(* IEC 61131-3 sources: Caravan/Archiv/12-04-19/Stations/Terminal/HMI/Class/_XMLReader (part 2) *)

  TextLen := _strlen(pText);
  TextLen += 1; // zero termination

  pDest^.pText$^void := StdLib.Malloc(TextLen);
  if pDest^.pText = NIL then
    XmlState := _ERROR;
    retcode := -2;
    return;
  end_if;

  _strcpy(pDest^.pText, pText);

  retcode := 0;

END_FUNCTION //AddTextAscii

FUNCTION _XMLReader::AddTextUni
	VAR_INPUT
		pDest 	: ^_XML_ELEMENT;
		pText 	: ^UINT;
	END_VAR
	VAR_OUTPUT
		retcode 	: DINT;
	END_VAR
  VAR
  	TextLen   : UDINT;
  END_VAR

  retcode := -1;

  if (pDest = NIL) | (pText = NIL) then
    return;
  end_if;

  // only allowed to add text when element has no children or already has a text
  if (pDest^.pText <> NIL) | (pDest^.pChildren <> NIL) then
    return;
  end_if;

  TextLen := SigCLib.StrLen16(pText)*2;
  TextLen += 2; // zero termination

  pDest^.pText$^void := StdLib.Malloc(TextLen);
  if pDest^.pText = NIL then
    XmlState := _ERROR;
    retcode := -2;
    return;
  end_if;

  SigCLib.StrCpy16(pDest^.pText$^UINT, pText);

  retcode := 0;

END_FUNCTION //AddTextUni

FUNCTION _XMLReader::CreateStructAscii
	VAR_INPUT
		parsedBytes 	: ^UDINT;
	END_VAR
	VAR_OUTPUT
		retcode 	: BOOL;
	END_VAR
VAR
	strBuff     : ^USINT;   // first tmp-Buffer
	strBuff2    : ^USINT;   // second tmp-Buffer
  pRun        : ^USINT;   // pointer to go through the information we read
  pStart      : ^USINT;   // points to the start of an element-name, atrib-name, attrib-value and so on...
  signCount   : UDINT;    // counts how much signs a string has
  counter     : UDINT;    // counter how far we passed through the information
  bufferLen   : UDINT;    // size of first buffer
  bufferLen2  : UDINT;    // size of second Buffer
END_VAR

  retcode := FALSE;

  // biggest work will be here
  // we have to go through the buffer and create our XML_STRUCT out of the information
  pRun := pFileBuffer;

  // set start size of buffer to 200, so in most cases we aren't going to resize the buffer
  // (normally names, values aren't this size, maybe text will be longer)
  bufferLen := 200;
  bufferLen2 := 200;

  strBuff$^void := StdLib.Malloc(bufferLen+1);
  strBuff2$^void := StdLib.Malloc(bufferLen2+1);

  if (strBuff = NIL) | (strBuff2 = NIL) then
    XmlState := _ERROR;
    return;
  end_if;

  _memset(strBuff, 0, bufferLen);
  _memset(strBuff2, 0, bufferLen2);

  counter := 1;

  // first handle the header
  if (pRun^ = XML_START) & ((pRun+1)^ = '?') then

    pStart := pRun;
    signCount := 0;

    while pRun^ <> XML_END do
      signCount += 1;

      counter += 1;
      pRun += 1;
    end_while;

    // now we are pointing at the end-mark, this also has to be in the header -> increase counters
    counter += 1;
    signCount += 1;

    if signCount > XML_MAX_HEADER_LENGTH then
      return;
    end_if;

    xmlStruct.Header$^void := StdLib.Malloc(signCount+1);
    _memset(xmlStruct.Header, 0, signCount+1);
    _memcpy(xmlStruct.Header, pStart, signCount);

    // alloc memory for first element and set struct for creator
    xmlStruct.MajorElement$^void := StdLib.Malloc(sizeof(_XML_ELEMENT));
    if (xmlStruct.MajorElement = NIL) then
      XmlState := _ERROR;
      return;
    end_if;
    _memset(xmlStruct.MajorElement, 0, sizeof(_XML_ELEMENT));
    StructCreator.SetStructPtr(#xmlStruct);

  else
    // xml does not start with the header
    ErrorState := _PARSE_ERR_NO_HEADER;
    parsedBytes^ := counter;
    return;
  end_if;

  // now lets see if we find a CR or LF and no signs between except of SPACE
  counter += 1;
  pRun += 1;
  while (pRun^ <> XML_CR) & (pRun^ <> XML_LF) do

    if pRun^ <> XML_SPACE then
      ErrorState := _PARSE_ERR_UNEXPECTED_SIGN;
      parsedBytes^ := counter;
      return; //wrong sign
    end_if;

    counter += 1;
    pRun += 1;
  end_while;

  // Header finished -> now lets start with looking for an Element
  searchFor := _SEARCH_ELEMENT;

  while counter < fileLength do

    case searchFor of

    	_SEARCH_ELEMENT:
    	  // look for '<'
        while pRun^ <> XML_START do

          if (pRun^ <> XML_CR) & (pRun^ <> XML_LF) & (pRun^ <> XML_SPACE) & (pRun^ <> XML_TABULATOR) then
            ErrorState := _PARSE_ERR_UNEXPECTED_SIGN;
            parsedBytes^ := counter;
            return; //wrong sign
          end_if;

          pRun += 1;
          counter += 1;
        end_while;

        // now we are pointing at start-mark, but we need one increase more
        pRun += 1;
        counter += 1;

        if (pRun^ <> XML_SLASH) & (pRun^ <> XML_EXCLAMATION) then
          //START Element
          if bTextSearched = TRUE then
            ErrorState := _PARSE_ERR_UNEXPECTED_SIGN;
            parsedBytes^ := counter;
            return; //wrong sign
          end_if;

          pStart := pRun;
          signCount := 0;

          // next step is to look for Space or End-Mark
          // counter are always one behind the pointer so we do not need to decrease afterwards
          while (pRun^ <> XML_END) & (pRun^ <> XML_SPACE) & (pRun^ <> XML_SLASH) do
            signCount += 1;

            counter += 1;
            pRun += 1;
          end_while;

          // at this point we found an element and we can get the name, so kick off name and add element to struct
          if signCount > bufferLen then
            bufferLen := signCount;
            StdLib.Free(strBuff);

            strBuff$^void := StdLib.Malloc(bufferLen+1);

            if (strBuff = NIL) then
              XmlState := _ERROR;
              return;
            end_if;

          end_if;

          _memcpy(strBuff, pStart, signCount);
          (strBuff+signCount)^ := 0;

          StructCreator.AddElement(strBuff, FALSE);

          // lets see what we have to do next
          if pRun^ = XML_END then

            pRun += 1;
            counter += 1;

            if (pRun^ = XML_CR) | (pRun^ = XML_LF) | (pRun^ = XML_START) | (pRun^ = XML_SPACE) then
              searchFor := _SEARCH_ELEMENT;
            else
              searchFor := _SEARCH_TEXT;
            end_if;

          elsif pRun^ = XML_SLASH then
            StructCreator.CloseElement(NIL,FALSE);

            // element is closed directly -> check if next sign is END-Tag
            pRun += 1;
            counter += 1;

            if pRun^ <> XML_END then
              // no end-tag after slash -> error
              ErrorState := _PARSE_ERR_UNEXPECTED_SIGN;
              parsedBytes^ := counter;
              return; //wrong sign
            end_if;

            // set to next sign
            pRun += 1;
            counter += 1;

            searchFor := _SEARCH_ELEMENT;

          elsif pRun^ = XML_SPACE then
            // in this case there can also be a closing-tag if element ist closed directly
            if (pRun+1)^ = XML_SLASH then

              StructCreator.CloseElement(NIL, FALSE);

              //                      <Element />
              //we point now to the space-----^---
              //but we need to be after end------^
              //this means +3 signs
              pRun += 3;
              counter += 3;

              searchFor := _SEARCH_ELEMENT;
            else
              searchFor := _SEARCH_ATTRIB;
            end_if;

          end_if;

        else
          if pRun^ = XML_SLASH then

            bTextSearched := FALSE;
            // CLOSE Element
            // so just go to the end of the close-element-tag and then close
            pRun += 1;
            counter += 1;

            pStart := pRun;
            signCount := 0;

            while pRun^ <> XML_END do
              signCount += 1;

              counter += 1;
              pRun += 1;
            end_while;

            if signCount > bufferLen then
              bufferLen := signCount;
              StdLib.Free(strBuff);

              strBuff$^void := StdLib.Malloc(bufferLen+1);
              if (strBuff = NIL) then
                XmlState := _ERROR;
                return;
              end_if;
            end_if;

            _memcpy(strBuff, pStart, signCount);
            (strBuff+signCount)^ := 0;

            pRun += 1;
            counter += 1;

            retClose := StructCreator.CloseElement(strBuff, FALSE);
            if retClose <> 0 then
              ErrorState := _PARSE_ERR_WRONG_SEQUENCE;
              parsedBytes^ := counter - signCount - 1;
              return; //wrong sequence of elements
            end_if;

            searchFor := _SEARCH_ELEMENT;

          else
            // check 4 comment
            if bTextSearched = TRUE then
              ErrorState := _PARSE_ERR_UNEXPECTED_SIGN;
              parsedBytes^ := counter;
              return; //wrong sign
            end_if;

            pRun += 1;
            counter += 1;
            if (pRun^ = XML_HYPHEN) & ((pRun+1)^ = XML_HYPHEN) then
              // we found '<!--' this means comment -> skip
              pRun += 2;
              counter += 2;

              while (pRun^ <> XML_HYPHEN) & ((pRun+1)^ <> XML_HYPHEN) & ((pRun+2)^ <> XML_END) do

                pRun += 1;
                counter += 1;

              end_while;
              pRun += 3; // set ptr to one ofter end-tag
              counter += 3;
              // we found the end '-->'
              // go on with searching for an element
              searchFor := _SEARCH_ELEMENT;

            end_if;

          end_if;

        end_if;

      _SEARCH_ATTRIB:

        bTextSearched := FALSE;
    	  // when we have to search 4 an attribute we know that pRun points to a Space
        // so the next sign is the start
        pRun += 1;
        counter += 1;

        pStart := pRun;
        signCount := 0;

        while pRun^ <> XML_EQUAL do

          if (pRun^ = XML_SPACE) | (pRun^ = XML_LF) | (pRun^ = XML_CR) then
            ErrorState := _PARSE_ERR_UNEXPECTED_SIGN;
            parsedBytes^ := counter;
            return; //wrong sign
          end_if;

          signCount += 1;
          counter += 1;
          pRun += 1;
        end_while;

        if signCount > bufferLen then
          bufferLen := signCount;
          StdLib.Free(strBuff);

          strBuff$^void := StdLib.Malloc(bufferLen+1);

          if (strBuff = NIL) then
            XmlState := _ERROR;
            return;
          end_if;

        end_if;

        _memcpy(strBuff, pStart, signCount);
        (strBuff+signCount)^ := 0;

        // we got the name of the attribute now lets get the value

        if ((pRun+1)^ <> XML_QUOTMARK) & ((pRun+1)^ <> XML_APOSTROPHE) then
          ErrorState := _PARSE_ERR_UNEXPECTED_SIGN;
          parsedBytes^ := counter;
          return; // wrong sign
        end_if;

        if ((pRun+1)^ = XML_QUOTMARK) then
          bQuot := TRUE;
        else
          bQuot := FALSE;
        end_if;

        pRun += 2; // set to one after quotation-mark
        counter += 2;

        pStart := pRun;
        signCount := 0;

        while ((pRun^ <> XML_QUOTMARK) & (bQuot = TRUE)) | ((pRun^ <> XML_APOSTROPHE) & (bQuot = FALSE)) do
          signCount += 1;

          counter += 1;
          pRun += 1;
        end_while;

        if signCount > bufferLen2 then
          bufferLen2 := signCount;
          StdLib.Free(strBuff2);

          strBuff2$^void := StdLib.Malloc(bufferLen2+1);

          if (strBuff2 = NIL) then
            XmlState := _ERROR;
            return;
          end_if;

        end_if;

        _memcpy(strBuff2, pStart, signCount);
        (strBuff2+signCount)^ := 0;

        if StructCreator.AddAttribute(strBuff, strBuff2, FALSE) = -1 then
          ErrorState := _PARSE_ERR_ATTRIBUTE_TWICE;
          parsedBytes^ := counter - signCount - 1;
          return; // attribute already exists
        end_if;

        // lets see what we have to do next
        pRun += 1;
        counter += 1;

        if pRun^ = XML_END then
          // so in this case we can have Text afterwards or next thing is an element
          pRun += 1;
          counter += 1;

          if (pRun^ = XML_CR) | (pRun^ = XML_LF) | (pRun^ = XML_START) then
            searchFor := _SEARCH_ELEMENT;
          else
            searchFor := _SEARCH_TEXT;
          end_if;

        elsif pRun^ = XML_SLASH then
            StructCreator.CloseElement(NIL, FALSE);

            // jump one sign after "/>"
            pRun += 2;
            counter += 2;
            searchFor := _SEARCH_ELEMENT;

        elsif pRun^ = XML_SPACE then
          // another attribute
          searchFor := _SEARCH_ATTRIB;
        end_if;

      _SEARCH_TEXT:
        // we already point to the start of the text
        pStart := pRun;
        signCount := 0;

        while pRun^ <> XML_START do
          signCount += 1;

          counter += 1;
          pRun += 1;
        end_while;

        if signCount > bufferLen then
          bufferLen := signCount;
          StdLib.Free(strBuff);

          strBuff$^void := StdLib.Malloc(bufferLen+1);

          if (strBuff = NIL) then
            XmlState := _ERROR;
            return;
          end_if;
        end_if;

        // kick off text & add to actual element
        _memcpy(strBuff, pStart, signCount);
        (strBuff+signCount)^ := 0;

        StructCreator.AddText(strBuff, FALSE);

        //next step hast to be looking for an element
        bTextSearched := TRUE;
        searchFor := _SEARCH_ELEMENT;

    end_case;

  end_while;

  StdLib.Free(strBuff);
  StdLib.Free(strBuff2);

  retcode := TRUE;

END_FUNCTION //CreateStructAscii

FUNCTION _XMLReader::CreateStructUni
	VAR_INPUT
		parsedBytes 	: ^UDINT;
	END_VAR
	VAR_OUTPUT
		retcode 	: BOOL;
	END_VAR
  VAR
    strBuff     : ^USINT;   // first tmp-Buffer
    strBuff2    : ^USINT;   // second tmp-Buffer
    pRun        : ^USINT;   // pointer to go through the information we read
    pStart      : ^USINT;   // points to the start of an element-name, atrib-name, attrib-value and so on...
    signCount   : UDINT;    // counts how much signs a string has
    counter     : UDINT;    // counter how far we passed through the information
    bufferLen   : UDINT;    // size of first buffer
    bufferLen2  : UDINT;    // size of second Buffer
  END_VAR

  retcode := FALSE;

  // biggest work will be here
  // we have to go through the buffer and create our XML_STRUCT out of the information
  pRun := pFileBuffer + 2;

  // set start size of buffer to 200, so in most cases we aren't going to resize the buffer
  // (normally names, values aren't this size, maybe text will be longer)
  bufferLen := 200;
  bufferLen2 := 200;

  strBuff$^void := StdLib.Malloc(bufferLen+2);
  strBuff2$^void := StdLib.Malloc(bufferLen2+2);

  if (strBuff = NIL) | (strBuff2 = NIL) then
    XmlState := _ERROR;
    return;
  end_if;

  _memset(strBuff, 0, bufferLen);
  _memset(strBuff2, 0, bufferLen2);

  counter := 2;

  // first handle the header
  if (pRun^$UINT = XML_START_UNI) & ((pRun+2)^$UINT = 16#003F) then

    pStart := pRun;
    signCount := 0;

    while pRun^$UINT <> XML_END_UNI do
      signCount += 2;

      counter += 2;
      pRun += 2;
    end_while;

    // now we are pointing at the end-mark, this also has to be in the header -> increase counters
    counter += 2;
    signCount += 2;

    if signCount > XML_MAX_HEADER_LENGTH then
      return;
    end_if;

    xmlStruct.Header$^void := StdLib.Malloc(signCount+2);
    _memset(xmlStruct.Header, 0, signCount+2);
    _memcpy(xmlStruct.Header, pStart, signCount);

    // alloc memory for first element and set struct for creator
    xmlStruct.MajorElement$^void := StdLib.Malloc(sizeof(_XML_ELEMENT));
    if (xmlStruct.MajorElement = NIL) then
      XmlState := _ERROR;
      return;
    end_if;
    _memset(xmlStruct.MajorElement, 0, sizeof(_XML_ELEMENT));
    StructCreator.SetStructPtr(#xmlStruct);

  else
    // xml does not start with the header
    ErrorState := _PARSE_ERR_NO_HEADER;
    parsedBytes^ := counter;
    return;
  end_if;

  // now lets see if we find a CR or LF and no signs between except of SPACE
  counter += 2;
  pRun += 2;
  while (pRun^$UINT <> XML_CR_UNI) & (pRun^$UINT <> XML_LF_UNI) do

    if pRun^$UINT <> XML_SPACE_UNI then
      ErrorState := _PARSE_ERR_UNEXPECTED_SIGN;
      parsedBytes^ := counter;
      return;
    end_if;

    counter += 2;
    pRun += 2;
  end_while;

  // Header finished -> now lets start with looking for an Element
  searchFor := _SEARCH_ELEMENT;

  while counter < fileLength do

    case searchFor of

    	_SEARCH_ELEMENT:
    	  // look for '<'
        while pRun^$UINT <> XML_START_UNI do

          if (pRun^$UINT <> XML_CR_UNI) & (pRun^$UINT <> XML_LF_UNI) & (pRun^$UINT <> XML_SPACE_UNI) & (pRun^$UINT <> XML_TABULATOR_UNI) then
            ErrorState := _PARSE_ERR_UNEXPECTED_SIGN;
            parsedBytes^ := counter;
            return;
          end_if;

          pRun += 2;
          counter += 2;
        end_while;

        // now we are pointing at start-mark, but we need one increase more
        pRun += 2;
        counter += 2;

        if (pRun^$UINT <> XML_SLASH_UNI) & (pRun^$UINT <> XML_EXCLAMATION_UNI) then
          //START Element
          if bTextSearched = TRUE then
            ErrorState := _PARSE_ERR_UNEXPECTED_SIGN;
            parsedBytes^ := counter;
            return;
          end_if;

          pStart := pRun;
          signCount := 0;

          // next step is to look for Space or End-Mark
          // counter are always one behind the pointer so we do not need to decrease afterwards
          while (pRun^$UINT <> XML_END_UNI) & (pRun^$UINT <> XML_SPACE_UNI) & (pRun^$UINT <> XML_SLASH_UNI) do
            signCount += 2;

            counter += 2;
            pRun += 2;
          end_while;

          // at this point we found an element and we can get the name, so kick off name and add element to struct
          if signCount > bufferLen then
            bufferLen := signCount;
            StdLib.Free(strBuff);

            strBuff$^void := StdLib.Malloc(bufferLen+2);

            if (strBuff = NIL) then
              XmlState := _ERROR;
              return;
            end_if;

          end_if;

          _memcpy(strBuff, pStart, signCount);
          (strBuff+signCount)^ := 0;
          (strBuff+signCount+1)^ := 0;

          StructCreator.AddElement(strBuff, TRUE);

          // lets see what we have to do next
          if pRun^$UINT = XML_END_UNI then

            pRun += 2;
            counter += 2;

            if (pRun^$UINT = XML_CR_UNI) | (pRun^$UINT = XML_LF_UNI) | (pRun^$UINT = XML_START_UNI) | (pRun^$UINT = XML_SPACE_UNI) then
              searchFor := _SEARCH_ELEMENT;
            else
              searchFor := _SEARCH_TEXT;
            end_if;

          elsif pRun^$UINT = XML_SLASH_UNI then
            StructCreator.CloseElement(NIL, TRUE);

            // element is closed directly -> check if next sign is END-Tag
            pRun += 2;
            counter += 2;

            if pRun^ <> XML_END_UNI then
              // no end-tag after slash -> error
              ErrorState := _PARSE_ERR_UNEXPECTED_SIGN;
              parsedBytes^ := counter;
              return;
            end_if;

            // set to next sign
            pRun += 2;
            counter += 2;

            searchFor := _SEARCH_ELEMENT;

          elsif pRun^$UINT = XML_SPACE_UNI then
            // in this case there can also be a closing-tag if element ist closed directly
            if (pRun+2)^ = XML_SLASH_UNI then

              StructCreator.CloseElement(NIL, TRUE);

              //                      <Element />
              //we point now to the space-----^---
              //but we need to be after end------^
              //this means +3 signs (in case of unicode 6Bytes)
              pRun += 6;
              counter += 6;

              searchFor := _SEARCH_ELEMENT;
            else
              searchFor := _SEARCH_ATTRIB;
            end_if;
          end_if;

        else
          if pRun^$UINT = XML_SLASH_UNI then

            bTextSearched := FALSE;
            // CLOSE Element
            // so just go to the end of the close-element-tag and then close
            pRun += 2;
            counter += 2;

            pStart := pRun;
            signCount := 0;

            while pRun^$UINT <> XML_END_UNI do
              signCount += 2;

              counter += 2;
              pRun += 2;
            end_while;

            if signCount > bufferLen then
              bufferLen := signCount;
              StdLib.Free(strBuff);
              strBuff$^void := StdLib.Malloc(bufferLen+2);
              if (strBuff = NIL) then
                XmlState := _ERROR;
                return;
              end_if;
            end_if;

            _memcpy(strBuff, pStart, signCount);
            (strBuff+signCount)^ := 0;
            (strBuff+signCount+1)^ := 0;
            pRun += 2;
            counter += 2;

            retClose := StructCreator.CloseElement(strBuff, TRUE);
            if retClose <> 0 then
              ErrorState := _PARSE_ERR_WRONG_SEQUENCE;
              parsedBytes^ := counter - signCount - 2;
              return;
            end_if;

            searchFor := _SEARCH_ELEMENT;

          else
            // check 4 comment
            if bTextSearched = TRUE then
              ErrorState := _PARSE_ERR_UNEXPECTED_SIGN;
              parsedBytes^ := counter;
              return;
            end_if;

            pRun += 2;
            counter += 2;
            if (pRun^$UINT = XML_HYPHEN_UNI) & ((pRun+1)^$UINT = XML_HYPHEN_UNI) then
              // we found '<!--' this means comment -> skip
              pRun += 4;
              counter += 4;

              while (pRun^$UINT <> XML_HYPHEN_UNI) & ((pRun+2)^$UINT <> XML_HYPHEN_UNI) & ((pRun+4)^$UINT <> XML_END_UNI) do

                pRun += 2;
                counter += 2;

              end_while;
              pRun += 6; // set ptr to one ofter end-tag
              counter += 6;
              // we found the end '-->'
              // go on with searching for an element
              searchFor := _SEARCH_ELEMENT;

            end_if;

          end_if;

        end_if;

      _SEARCH_ATTRIB:

        bTextSearched := FALSE;
    	  // when we have to search 4 an attribute we know that pRun points to a Space
        // so the next sign is the start
        pRun += 2;
        counter += 2;

        pStart := pRun;
        signCount := 0;

        while pRun^$UINT <> XML_EQUAL_UNI do

          if (pRun^$UINT = XML_SPACE_UNI) | (pRun^$UINT = XML_LF_UNI) | (pRun^$UINT = XML_CR_UNI) then
            ErrorState := _PARSE_ERR_UNEXPECTED_SIGN;
            parsedBytes^ := counter;
            return;
          end_if;

          signCount += 2;
          counter += 2;
          pRun += 2;
        end_while;

        if signCount > bufferLen then
          bufferLen := signCount;
          StdLib.Free(strBuff);

          strBuff$^void := StdLib.Malloc(bufferLen+2);

          if (strBuff = NIL) then
            XmlState := _ERROR;
            return;
          end_if;

        end_if;

        _memcpy(strBuff, pStart, signCount);
        (strBuff+signCount)^ := 0;
        (strBuff+signCount+1)^ := 0;

        // we got the name of the attribute now lets get the value

        if ((pRun+2)^$UINT <> XML_QUOTMARK_UNI) & ((pRun+2)^$UINT <> XML_APOSTROPHE_UNI) then
          ErrorState := _PARSE_ERR_UNEXPECTED_SIGN;
          parsedBytes^ := counter;
          return;
        end_if;

        if ((pRun+2)^$UINT = XML_QUOTMARK_UNI) then
          bQuot := TRUE;
        else
          bQuot := FALSE;
        end_if;

        pRun += 4; // set to one after quotation-mark
        counter += 4;

        pStart := pRun;
        signCount := 0;

        while ((pRun^$UINT <> XML_QUOTMARK_UNI) & (bQuot = TRUE)) | ((pRun^$UINT <> XML_APOSTROPHE_UNI) & (bQuot = FALSE)) do
          signCount += 2;

          counter += 2;
          pRun += 2;
        end_while;

        if signCount > bufferLen2 then
          bufferLen2 := signCount;
          StdLib.Free(strBuff2);
          strBuff2$^void := StdLib.Malloc(bufferLen2+2);

          if (strBuff2 = NIL) then
            XmlState := _ERROR;
            return;
          end_if;

        end_if;

        _memcpy(strBuff2, pStart, signCount);
        (strBuff2+signCount)^ := 0;
        (strBuff2+signCount + 1)^ := 0;
        if StructCreator.AddAttribute(strBuff, strBuff2, TRUE) = -1 then
          ErrorState := _PARSE_ERR_ATTRIBUTE_TWICE;
          parsedBytes^ := counter - signCount - 2;
          return; // attribute already exists
        end_if;

        // lets see what we have to do next
        pRun += 2;
        counter += 2;

        if pRun^$UINT = XML_END_UNI then
          // so in this case we can have Text afterwards or next thing is an element
          pRun += 2;
          counter += 2;

          if (pRun^$UINT = XML_CR_UNI) | (pRun^$UINT = XML_LF_UNI) | (pRun^$UINT = XML_START_UNI) then
            searchFor := _SEARCH_ELEMENT;
          else
            searchFor := _SEARCH_TEXT;
          end_if;

        elsif pRun^$UINT = XML_SLASH_UNI then
            StructCreator.CloseElement(NIL, TRUE);

            // jump one sign after "/>"
            pRun += 4;
            counter += 4;
            searchFor := _SEARCH_ELEMENT;

        elsif pRun^$UINT = XML_SPACE_UNI then
          // another attribute
          searchFor := _SEARCH_ATTRIB;
        end_if;

      _SEARCH_TEXT:
        // we already point to the start of the text
        pStart := pRun;
        signCount := 0;

        while pRun^$UINT <> XML_START_UNI do
          signCount += 2;

          counter += 2;
          pRun += 2;
        end_while;

        if signCount > bufferLen then
          bufferLen := signCount;
          StdLib.Free(strBuff);

          strBuff$^void := StdLib.Malloc(bufferLen+2);

          if (strBuff = NIL) then
            XmlState := _ERROR;
            return;
          end_if;
        end_if;

        // kick off text & add to actual element
        _memcpy(strBuff, pStart, signCount);
        (strBuff+signCount)^ := 0;
        (strBuff+signCount + 1)^ := 0;
        StructCreator.AddText(strBuff, TRUE);

        //next step hast to be looking for an element
        bTextSearched := TRUE;
        searchFor := _SEARCH_ELEMENT;

    end_case;

  end_while;

  StdLib.Free(strBuff);
  StdLib.Free(strBuff2);

  retcode := TRUE;

END_FUNCTION //CreateStructUni

FUNCTION _XMLReader::FindError
	VAR_INPUT
		bytesParsed 	: UDINT;
	END_VAR
  VAR
  	count : UDINT;
    linecount : UDINT;
    signsUntilCRLF : UDINT;
    pTmp  : ^USINT;
  END_VAR

  lineCount := 1;
  signsUntilCRLF := 0;

  pTmp := pFileBuffer;

  if bRdIsUnicode = TRUE then
    pTmp += sizeof(UINT);

    bytesParsed := bytesParsed / 2;
  end_if;

  for count := 1 to bytesParsed - 1 do

    if pTmp^ = XML_LF | pTmp^ = XML_CR then
      linecount += 1;
      signsUntilCRLF := 0;

      while pTmp^ = XML_CR | pTmp^ = XML_LF do
        if bRdIsUnicode = TRUE then
          pTmp += sizeof(UINT);
        else
          pTmp += sizeof(USINT);
        end_if;
      end_while;

    else
      signsUntilCRLF += 1;

      if bRdIsUnicode = TRUE then
        pTmp += sizeof(UINT);
      else
        pTmp += sizeof(USINT);
      end_if;
    end_if;

  end_for;

  ErrorLine := TO_DINT(linecount);
  ErrorSign := TO_DINT(signsUntilCRLF);

END_FUNCTION

FUNCTION GLOBAL _XMLReader::GetAttribValueByName
	VAR_INPUT
		pElement 	: ^_XML_ELEMENT;
		pName 	: ^USINT;
	END_VAR
	VAR_OUTPUT
		pValue 	: ^USINT;
	END_VAR

  if pElement = NIL | pName = NIL then
    pValue := NIL;
    return;
  end_if;

  // look if we have tu use unicode functions or not
  if bRdIsUnicode = TRUE then
    pValue := GetAttribValueByNameUni(pElement, pName$^UINT);
  else
    pValue := GetAttribValueByNameAscii(pElement, pName);
  end_if;

END_FUNCTION

FUNCTION _XMLReader::GetAttribValueByNameAscii
	VAR_INPUT
		pElement 	: ^_XML_ELEMENT;
		pName 	: ^USINT;
	END_VAR
	VAR_OUTPUT
		pValue 	: ^USINT;
	END_VAR
  VAR
  	i : UDINT;
    pAttrib : ^_XML_ATTRIBUTE;
  END_VAR

  pValue := NIL;

  // go through whole attribute list and check names
  pAttrib := pElement^.Attributes.pList;
  for i := 1 to pElement^.Attributes.no do

    if SigCLib.StrCmp(pName, pAttrib^.Name) = 0 then
      pValue := pAttrib^.Value;
      return;
    end_if;

    pAttrib += sizeof(_XML_ATTRIBUTE);
  end_for;

END_FUNCTION

FUNCTION _XMLReader::GetAttribValueByNameUni
	VAR_INPUT
		pElement 	: ^_XML_ELEMENT;
		pName 	: ^UINT;
	END_VAR
	VAR_OUTPUT
		pValue 	: ^USINT;
	END_VAR
  VAR
  	i : UDINT;
    pAttrib : ^_XML_ATTRIBUTE;
  END_VAR

  pValue := NIL;

  // go through whole attribute list and check names
  pAttrib := pElement^.Attributes.pList;
  for i := 1 to pElement^.Attributes.no do

    if SigCLib.StrCmp16(pName, pAttrib^.Name$^UINT) = 0 then
      pValue := pAttrib^.Value;
      return;
    end_if;

    pAttrib += sizeof(_XML_ATTRIBUTE);
  end_for;

END_FUNCTION

FUNCTION GLOBAL _XMLReader::GetChildByName
	VAR_INPUT
		pParent 	: ^_XML_ELEMENT;
		pName 	: ^USINT;
		number 	: UDINT;(* := 1 *)
	END_VAR
	VAR_OUTPUT
		pChild 	: ^_XML_ELEMENT;
	END_VAR

  // number = 1 means first child; number = 2 means second child and so on...
  if number = 0 then
    pChild := NIL;
    return;
  end_if;

  if pParent = NIL | pName = NIL then
    pChild := NIL;
    return;
  end_if;

  if bRdIsUnicode = TRUE then
    pChild := GetChildByNameUni(pParent, pName$^UINT, number);
  else
    pChild := GetChildByNameAscii(pParent, pName, number);
  end_if;

END_FUNCTION

FUNCTION _XMLReader::GetChildByNameAscii
	VAR_INPUT
		pParent 	: ^_XML_ELEMENT;
		pName 	: ^USINT;
		number 	: UDINT;
	END_VAR
	VAR_OUTPUT
		pChild 	: ^_XML_ELEMENT;
	END_VAR
  VAR
  	pTmp : ^_XML_ELEMENT;
    tmpNr : UDINT;
  END_VAR

  pChild := NIL;

  // set temp-pointer to first child
  pTmp := pParent^.pChildren;
  tmpNr := number;

  while pTmp <> NIL do
    // go through childs and compare names
    if SigCLib.StrCmp(pTmp^.Name, pName) = 0 then

      tmpNr -= 1;
      if tmpNr = 0 then
        pChild := pTmp;
        return;
      end_if;

    end_if;

    pTmp := pTmp^.pNext;
  end_while;

END_FUNCTION

FUNCTION _XMLReader::GetChildByNameUni
	VAR_INPUT
		pParent 	: ^_XML_ELEMENT;
		pName 	: ^UINT;
		number 	: UDINT;
	END_VAR
	VAR_OUTPUT
		pChild 	: ^_XML_ELEMENT;
	END_VAR
  VAR
  	pTmp : ^_XML_ELEMENT;
    tmpNr : UDINT;
  END_VAR

  pChild := NIL;

  // set temp-pointer to first child
  pTmp := pParent^.pChildren;
  tmpNr := number;

  while pTmp <> NIL do
    // go through childs and compare names
    if SigCLib.StrCmp16(pTmp^.Name$^UINT, pName) = 0 then

      tmpNr -= 1;
      if tmpNr = 0 then
        pChild := pTmp;
        return;
      end_if;

    end_if;

    pTmp := pTmp^.pNext;
  end_while;

END_FUNCTION

FUNCTION GLOBAL _XMLReader::ParseXML
	VAR_INPUT
		pData 	: ^USINT;
		length 	: UDINT;
	END_VAR
	VAR_OUTPUT
		retcode 	: BOOL;
	END_VAR

  retcode := FALSE;

  if XmlState = _READY then // check if reader is ready

    if length > 0 then // check given length

      pFileBuffer$^void := StdLib.Malloc(length);
      if pFileBuffer <> NIL then

        // alloc memory was successfull - copy data
        _memcpy(pFileBuffer, pData, length);

        fileLength := length;

        XmlState := _PARSE_STREAM;
        readSSW := _CREATE_STRUCT;

        retcode := TRUE;
      end_if;

    end_if;

  end_if;

END_FUNCTION

FUNCTION GLOBAL _XMLReader::GetXmlState
	VAR_OUTPUT
		state 	: XML_READ_STATE;
	END_VAR

  state := XmlState;

END_FUNCTION

FUNCTION GLOBAL _XMLReader::GetErrorState
	VAR_OUTPUT
		state 	: _XML_PARSE_ERROR;
	END_VAR

  state := ErrorState;

END_FUNCTION
